// TIA Portal V21 export
// export: Created 2026-11-10T19:11:39.1091354Z, ExportSetting WithDefaults, DisplayName Totally Integrated Automation Portal, DisplayVersion V21 Update 3, DisplayName STEP 7 Professional, DisplayVersion V21 Update 3, DisplayName STEP 7 Safety, DisplayVersion V21, DisplayName Tech WebApplication, DisplayVersion V21, DisplayName WinCC Basic/Comfort/Advanced, DisplayVersion V21 Update 3, DisplayName WinCC Unified, DisplayVersion V21 Update 3
DATA_BLOCK "DB_PULSEGEN"   // DB28
// stored: AutoNumber true, DBAccessibleFromOPCUA true, DBAccessibleFromWebserver true, InstanceOfName PULSEGEN, OfSystemLibElement PULSEGEN, OfSystemLibVersion 1.1
"PULSEGEN"
   // VAR_INPUT
   //    INV : Real;
   //    PER_TM : Time;
   //    P_B_TM : Time;
   //    RATIOFAC : Real;
   //    STEP3_ON : Bool;
   //    ST2BI_ON : Bool;
   //    MAN_ON : Bool;
   //    POS_P_ON : Bool;
   //    NEG_P_ON : Bool;
   //    SYN_ON : Bool;
   //    COM_RST : Bool;
   //    CYCLE : Time;
   // END_VAR
   // VAR_OUTPUT
   //    QPOS_P : Bool;
   //    QNEG_P : Bool;
   // END_VAR
   // VAR RETAIN
   //    sInvAlt : Real;
   //    siZaehlPer : Int;
   //    siZaehlPTm : Int;
   //    sbPosP : Bool;
   // END_VAR
BEGIN
END_DATA_BLOCK
